(* IEC 61131-3 sources: Test-Git_ESME26/TestProgettoESME_26.fbsproj/PacDriveLib Migration/LibraryDiagnostics, 1 file *)

(* ---- PDL_FC_EtDiagExtToString.fn.st ---- *)
FUNCTION PDL_FC_EtDiagExtToString : STRING[80]
VAR_INPUT
	i_etDiagExt : PDL_ET_DiagExt;
END_VAR
VAR_OUTPUT
	q_etDiag			: GD.ET_Diag := GD.ET_Diag.OK;
	q_etDiagExt			: PDL_ET_DiagExt := PDL_ET_DiagExt.OK;
END_VAR
VAR
END_VAR

PDL_FC_EtDiagExtToString := TO_STRING(i_etDiagExt);
